Fanuc KAREL source: KO00112.KL

PROGRAM KO00112
%NOLOCKGROUP
VAR
  A: REAL
  B: ARRAY[2] OF SHORT
  OUT: REAL
BEGIN
  A = 1
  B[1] = 2
  OUT = ATAN2(A, B[1])
END KO00112
